// Mitsubishi GX Works2 project: SEMICON_SORTER_ENV   PLC: FX3U/FX3UC

PROGRAM MAIN
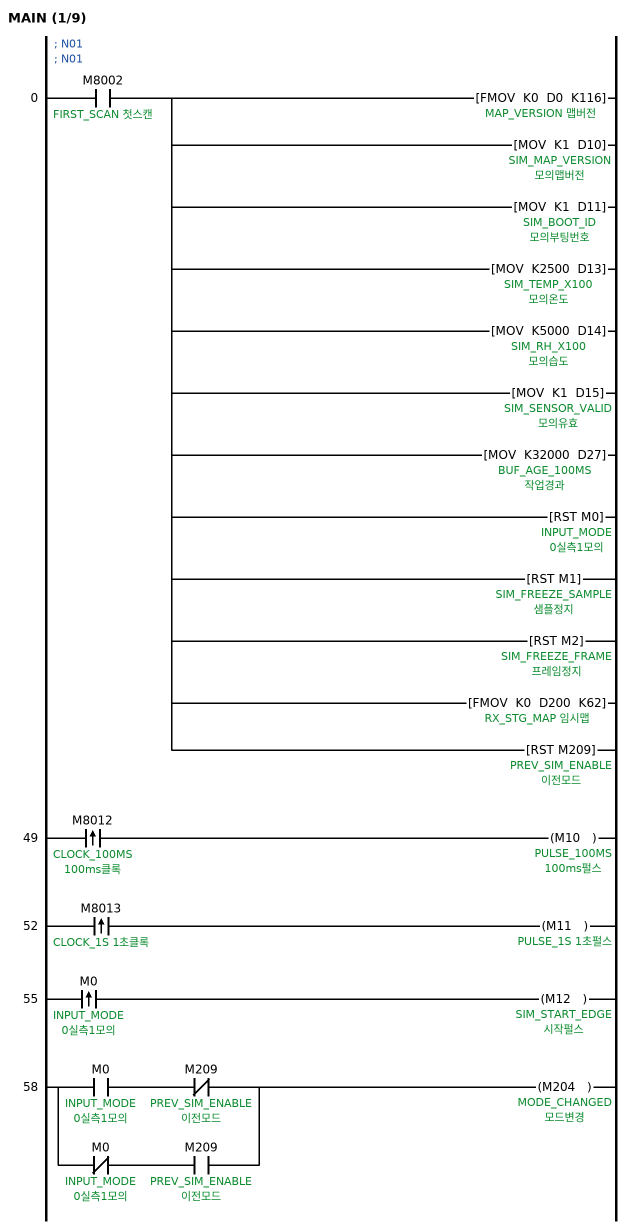
; 
; N01
; N01
0     LD      M8002  ; FIRST_SCAN 첫스캔
      FMOV    K0 D0 K116  ; MAP_VERSION 맵버전
      MOV     K1 D10  ; SIM_MAP_VERSION 모의맵버전
      MOV     K1 D11  ; SIM_BOOT_ID 모의부팅번호
      MOV     K2500 D13  ; SIM_TEMP_X100 모의온도
      MOV     K5000 D14  ; SIM_RH_X100 모의습도
      MOV     K1 D15  ; SIM_SENSOR_VALID 모의유효
      MOV     K32000 D27  ; BUF_AGE_100MS 작업경과
      RST     M0  ; INPUT_MODE 0실측1모의
      RST     M1  ; SIM_FREEZE_SAMPLE 샘플정지
      RST     M2  ; SIM_FREEZE_FRAME 프레임정지
      FMOV    K0 D200 K62  ; RX_STG_MAP 임시맵
      RST     M209  ; PREV_SIM_ENABLE 이전모드
49    LDP     M8012  ; CLOCK_100MS 100ms클록
      OUT     M10  ; PULSE_100MS 100ms펄스
52    LDP     M8013  ; CLOCK_1S 1초클록
      OUT     M11  ; PULSE_1S 1초펄스
55    LDP     M0  ; INPUT_MODE 0실측1모의
      OUT     M12  ; SIM_START_EDGE 시작펄스
58    LD      M0  ; INPUT_MODE 0실측1모의
      ANI     M209  ; PREV_SIM_ENABLE 이전모드
      LDI     M0  ; INPUT_MODE 0실측1모의
      AND     M209  ; PREV_SIM_ENABLE 이전모드
      ORB
      OUT     M204  ; MODE_CHANGED 모드변경
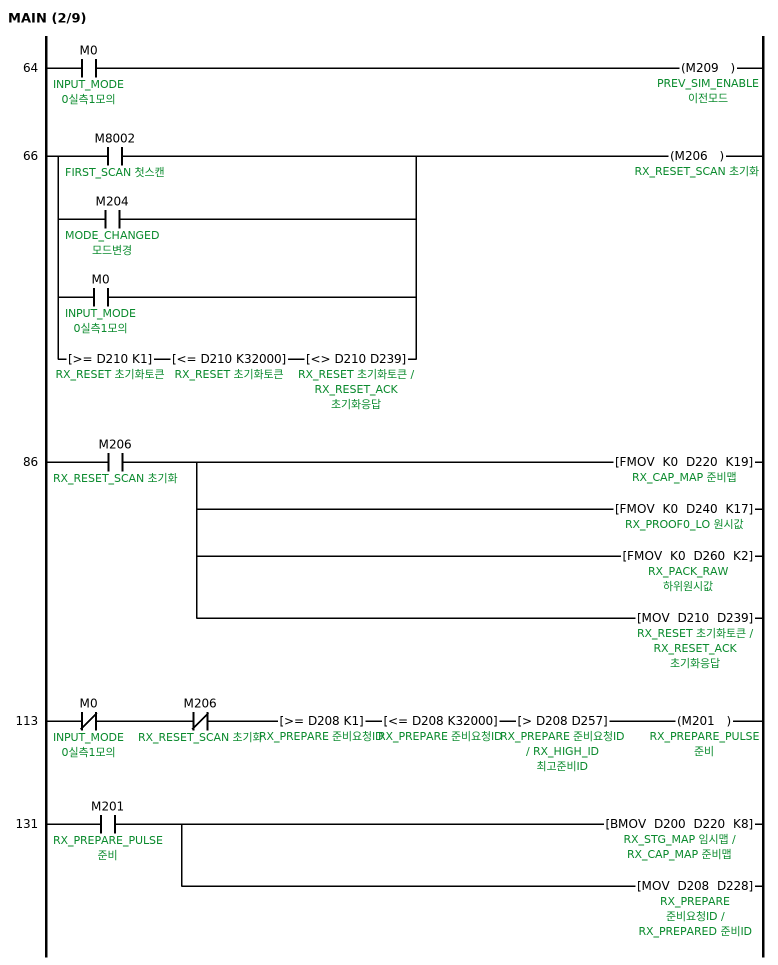
64    LD      M0  ; INPUT_MODE 0실측1모의
      OUT     M209  ; PREV_SIM_ENABLE 이전모드
66    LD      M8002  ; FIRST_SCAN 첫스캔
      OR      M204  ; MODE_CHANGED 모드변경
      OR      M0  ; INPUT_MODE 0실측1모의
      LD>=    D210 K1  ; RX_RESET 초기화토큰
      AND<=   D210 K32000  ; RX_RESET 초기화토큰
      AND<>   D210 D239  ; RX_RESET 초기화토큰 / RX_RESET_ACK 초기화응답
      ORB
      OUT     M206  ; RX_RESET_SCAN 초기화
86    LD      M206  ; RX_RESET_SCAN 초기화
      FMOV    K0 D220 K19  ; RX_CAP_MAP 준비맵
      FMOV    K0 D240 K17  ; RX_PROOF0_LO 원시값
      FMOV    K0 D260 K2  ; RX_PACK_RAW 하위원시값
      MOV     D210 D239
113   LDI     M0  ; INPUT_MODE 0실측1모의
      ANI     M206  ; RX_RESET_SCAN 초기화
      AND>=   D208 K1  ; RX_PREPARE 준비요청ID
      AND<=   D208 K32000  ; RX_PREPARE 준비요청ID
      AND>    D208 D257  ; RX_PREPARE 준비요청ID / RX_HIGH_ID 최고준비ID
      OUT     M201  ; RX_PREPARE_PULSE 준비
131   LD      M201  ; RX_PREPARE_PULSE 준비
      BMOV    D200 D220 K8
      MOV     D208 D228  ; RX_PREPARED 준비ID
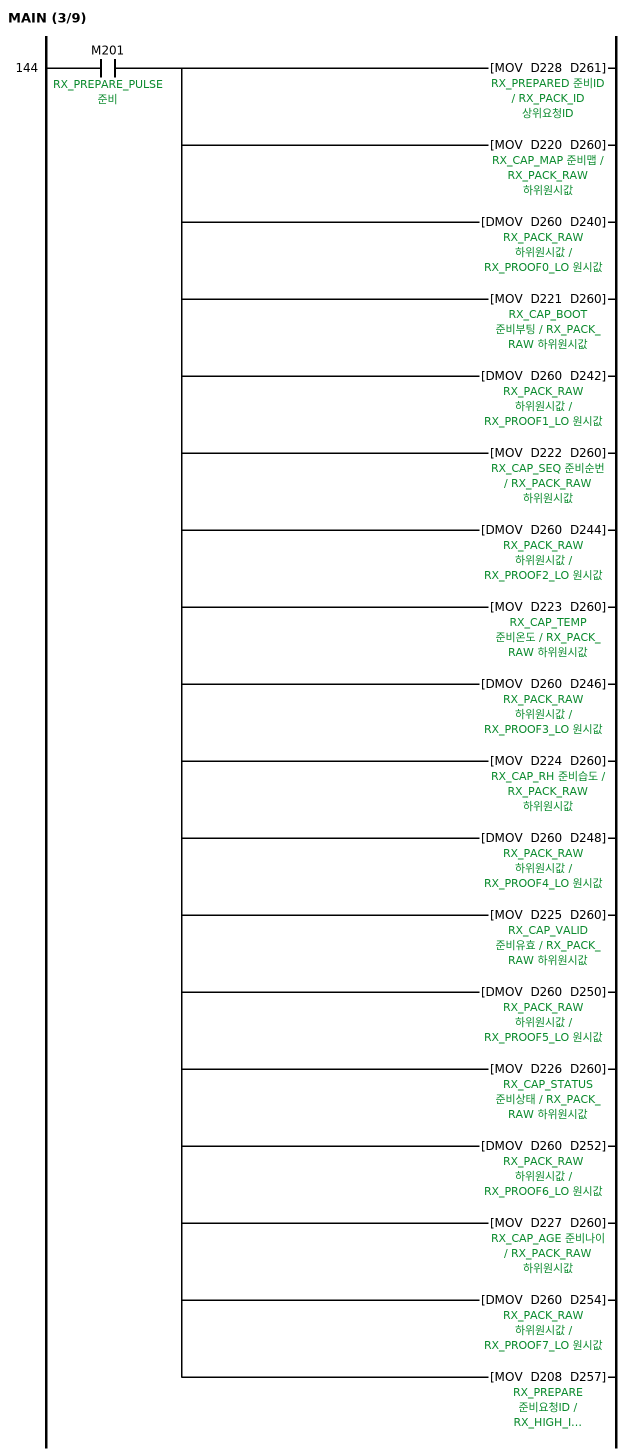
144   LD      M201  ; RX_PREPARE_PULSE 준비
      MOV     D228 D261  ; RX_PACK_ID 상위요청ID
      MOV     D220 D260
      DMOV    D260 D240
      MOV     D221 D260  ; RX_CAP_BOOT 준비부팅
      DMOV    D260 D242  ; RX_PROOF1_LO 원시값
      MOV     D222 D260  ; RX_CAP_SEQ 준비순번
      DMOV    D260 D244  ; RX_PROOF2_LO 원시값
      MOV     D223 D260  ; RX_CAP_TEMP 준비온도
      DMOV    D260 D246  ; RX_PROOF3_LO 원시값
      MOV     D224 D260  ; RX_CAP_RH 준비습도
      DMOV    D260 D248  ; RX_PROOF4_LO 원시값
      MOV     D225 D260  ; RX_CAP_VALID 준비유효
      DMOV    D260 D250  ; RX_PROOF5_LO 원시값
      MOV     D226 D260  ; RX_CAP_STATUS 준비상태
      DMOV    D260 D252  ; RX_PROOF6_LO 원시값
      MOV     D227 D260  ; RX_CAP_AGE 준비나이
      DMOV    D260 D254  ; RX_PROOF7_LO 원시값
      MOV     D208 D257
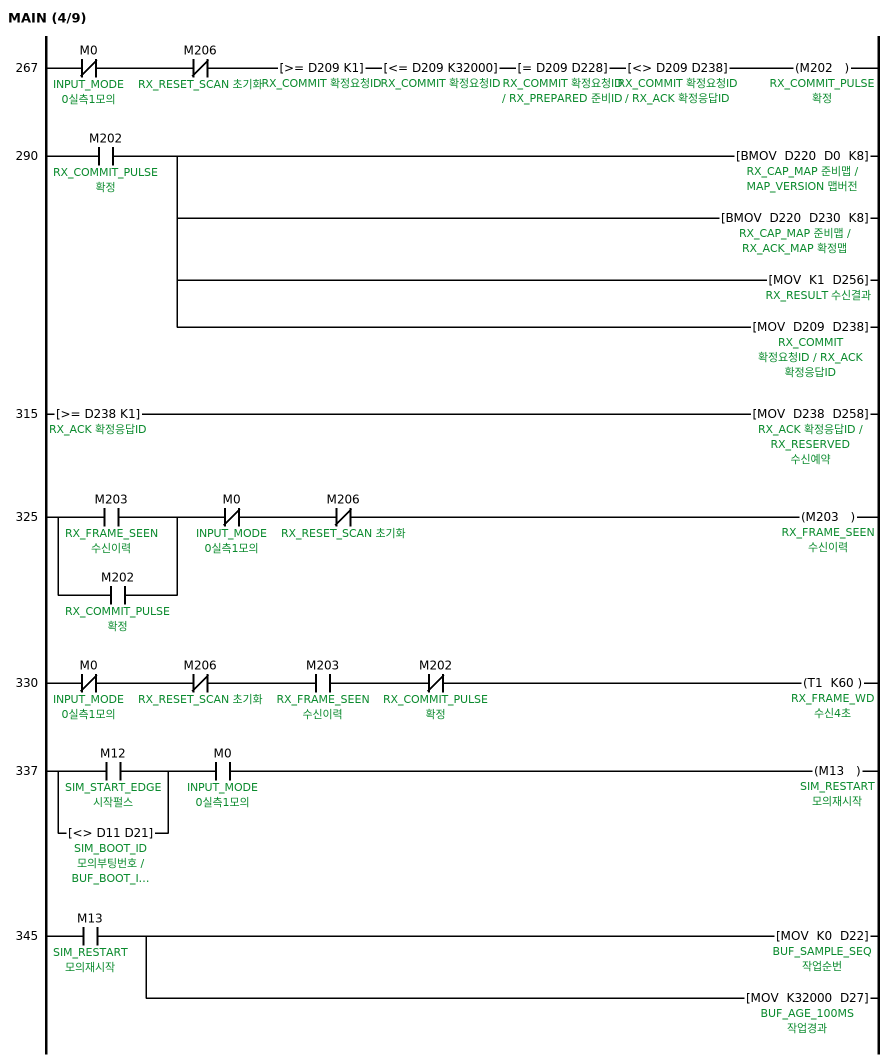
267   LDI     M0  ; INPUT_MODE 0실측1모의
      ANI     M206  ; RX_RESET_SCAN 초기화
      AND>=   D209 K1  ; RX_COMMIT 확정요청ID
      AND<=   D209 K32000  ; RX_COMMIT 확정요청ID
      AND=    D209 D228  ; RX_COMMIT 확정요청ID / RX_PREPARED 준비ID
      AND<>   D209 D238  ; RX_COMMIT 확정요청ID / RX_ACK 확정응답ID
      OUT     M202  ; RX_COMMIT_PULSE 확정
290   LD      M202  ; RX_COMMIT_PULSE 확정
      BMOV    D220 D0 K8
      BMOV    D220 D230 K8  ; RX_ACK_MAP 확정맵
      MOV     K1 D256  ; RX_RESULT 수신결과
      MOV     D209 D238
315   LD>=    D238 K1  ; RX_ACK 확정응답ID
      MOV     D238 D258  ; RX_RESERVED 수신예약
325   LD      M203  ; RX_FRAME_SEEN 수신이력
      OR      M202  ; RX_COMMIT_PULSE 확정
      ANI     M0  ; INPUT_MODE 0실측1모의
      ANI     M206  ; RX_RESET_SCAN 초기화
      OUT     M203  ; RX_FRAME_SEEN 수신이력
330   LDI     M0  ; INPUT_MODE 0실측1모의
      ANI     M206  ; RX_RESET_SCAN 초기화
      AND     M203  ; RX_FRAME_SEEN 수신이력
      ANI     M202  ; RX_COMMIT_PULSE 확정
      OUT     T1 K60  ; RX_FRAME_WD 수신4초
337   LD      M12  ; SIM_START_EDGE 시작펄스
      OR<>    D11 D21  ; SIM_BOOT_ID 모의부팅번호 / BUF_BOOT_ID 작업부팅번호
      AND     M0  ; INPUT_MODE 0실측1모의
      OUT     M13  ; SIM_RESTART 모의재시작
345   LD      M13  ; SIM_RESTART 모의재시작
      MOV     K0 D22  ; BUF_SAMPLE_SEQ 작업순번
      MOV     K32000 D27
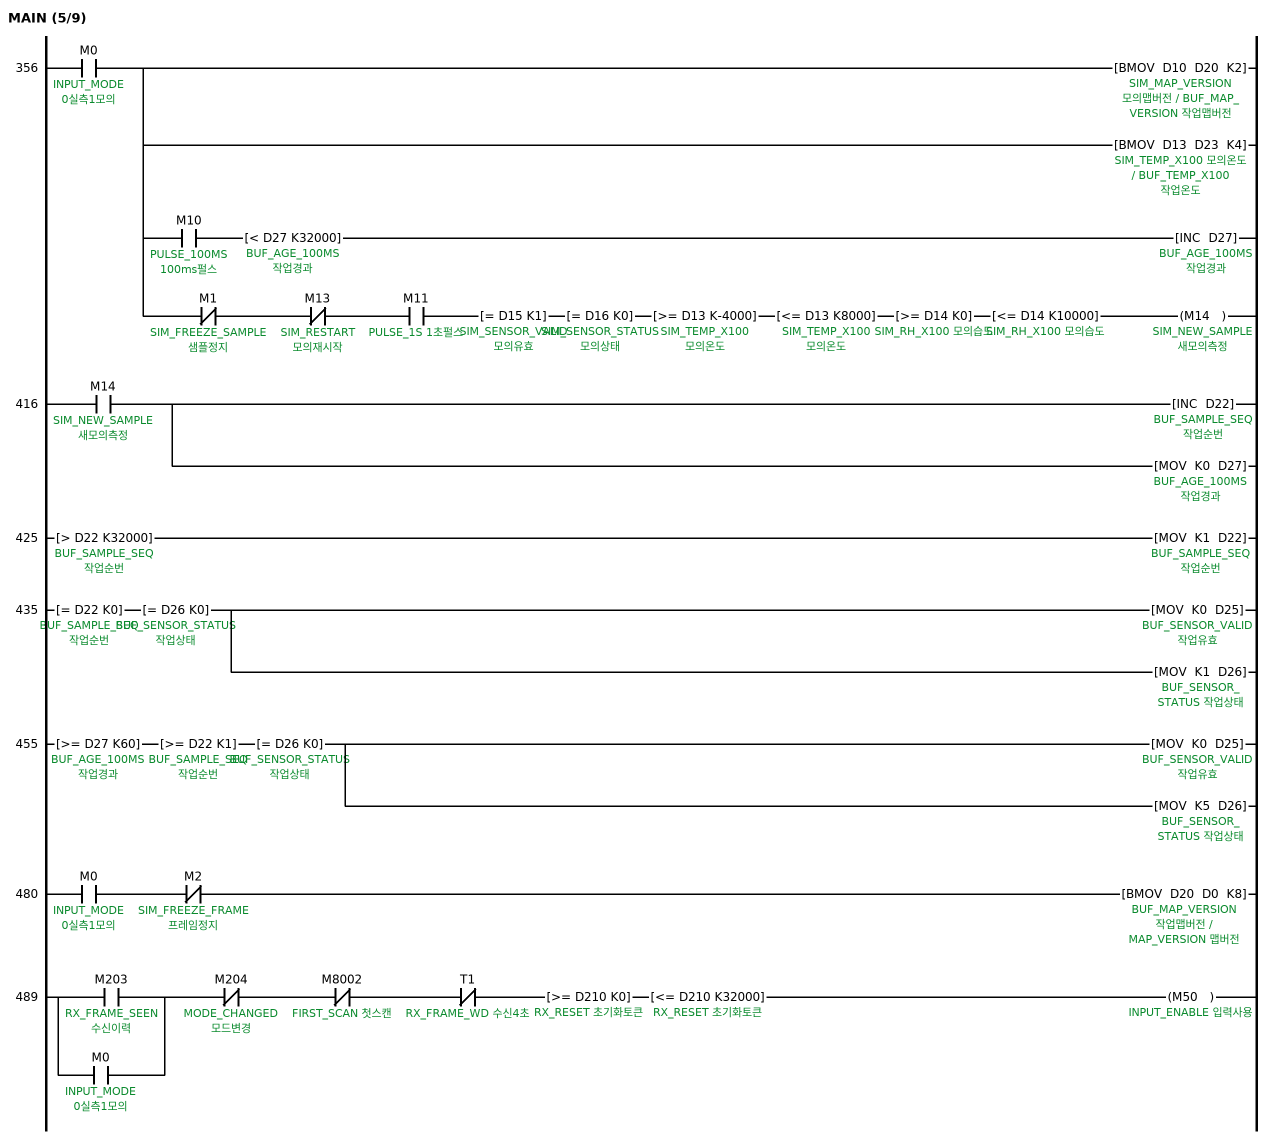
356   LD      M0  ; INPUT_MODE 0실측1모의
      BMOV    D10 D20 K2  ; BUF_MAP_VERSION 작업맵버전
      BMOV    D13 D23 K4  ; BUF_TEMP_X100 작업온도
      MPS
      AND     M10  ; PULSE_100MS 100ms펄스
      AND<    D27 K32000  ; BUF_AGE_100MS 작업경과
      INC     D27
      MPP
      ANI     M1  ; SIM_FREEZE_SAMPLE 샘플정지
      ANI     M13  ; SIM_RESTART 모의재시작
      AND     M11  ; PULSE_1S 1초펄스
      AND=    D15 K1  ; SIM_SENSOR_VALID 모의유효
      AND=    D16 K0  ; SIM_SENSOR_STATUS 모의상태
      AND>=   D13 K-4000  ; SIM_TEMP_X100 모의온도
      AND<=   D13 K8000  ; SIM_TEMP_X100 모의온도
      AND>=   D14 K0  ; SIM_RH_X100 모의습도
      AND<=   D14 K10000  ; SIM_RH_X100 모의습도
      OUT     M14  ; SIM_NEW_SAMPLE 새모의측정
416   LD      M14  ; SIM_NEW_SAMPLE 새모의측정
      INC     D22
      MOV     K0 D27
425   LD>     D22 K32000  ; BUF_SAMPLE_SEQ 작업순번
      MOV     K1 D22
435   LD=     D22 K0  ; BUF_SAMPLE_SEQ 작업순번
      AND=    D26 K0  ; BUF_SENSOR_STATUS 작업상태
      MOV     K0 D25  ; BUF_SENSOR_VALID 작업유효
      MOV     K1 D26
455   LD>=    D27 K60  ; BUF_AGE_100MS 작업경과
      AND>=   D22 K1  ; BUF_SAMPLE_SEQ 작업순번
      AND=    D26 K0  ; BUF_SENSOR_STATUS 작업상태
      MOV     K0 D25
      MOV     K5 D26
480   LD      M0  ; INPUT_MODE 0실측1모의
      ANI     M2  ; SIM_FREEZE_FRAME 프레임정지
      BMOV    D20 D0 K8
489   LD      M203  ; RX_FRAME_SEEN 수신이력
      OR      M0  ; INPUT_MODE 0실측1모의
      ANI     M204  ; MODE_CHANGED 모드변경
      ANI     M8002  ; FIRST_SCAN 첫스캔
      ANI     T1  ; RX_FRAME_WD 수신4초
      AND>=   D210 K0  ; RX_RESET 초기화토큰
      AND<=   D210 K32000  ; RX_RESET 초기화토큰
      OUT     M50  ; INPUT_ENABLE 입력사용
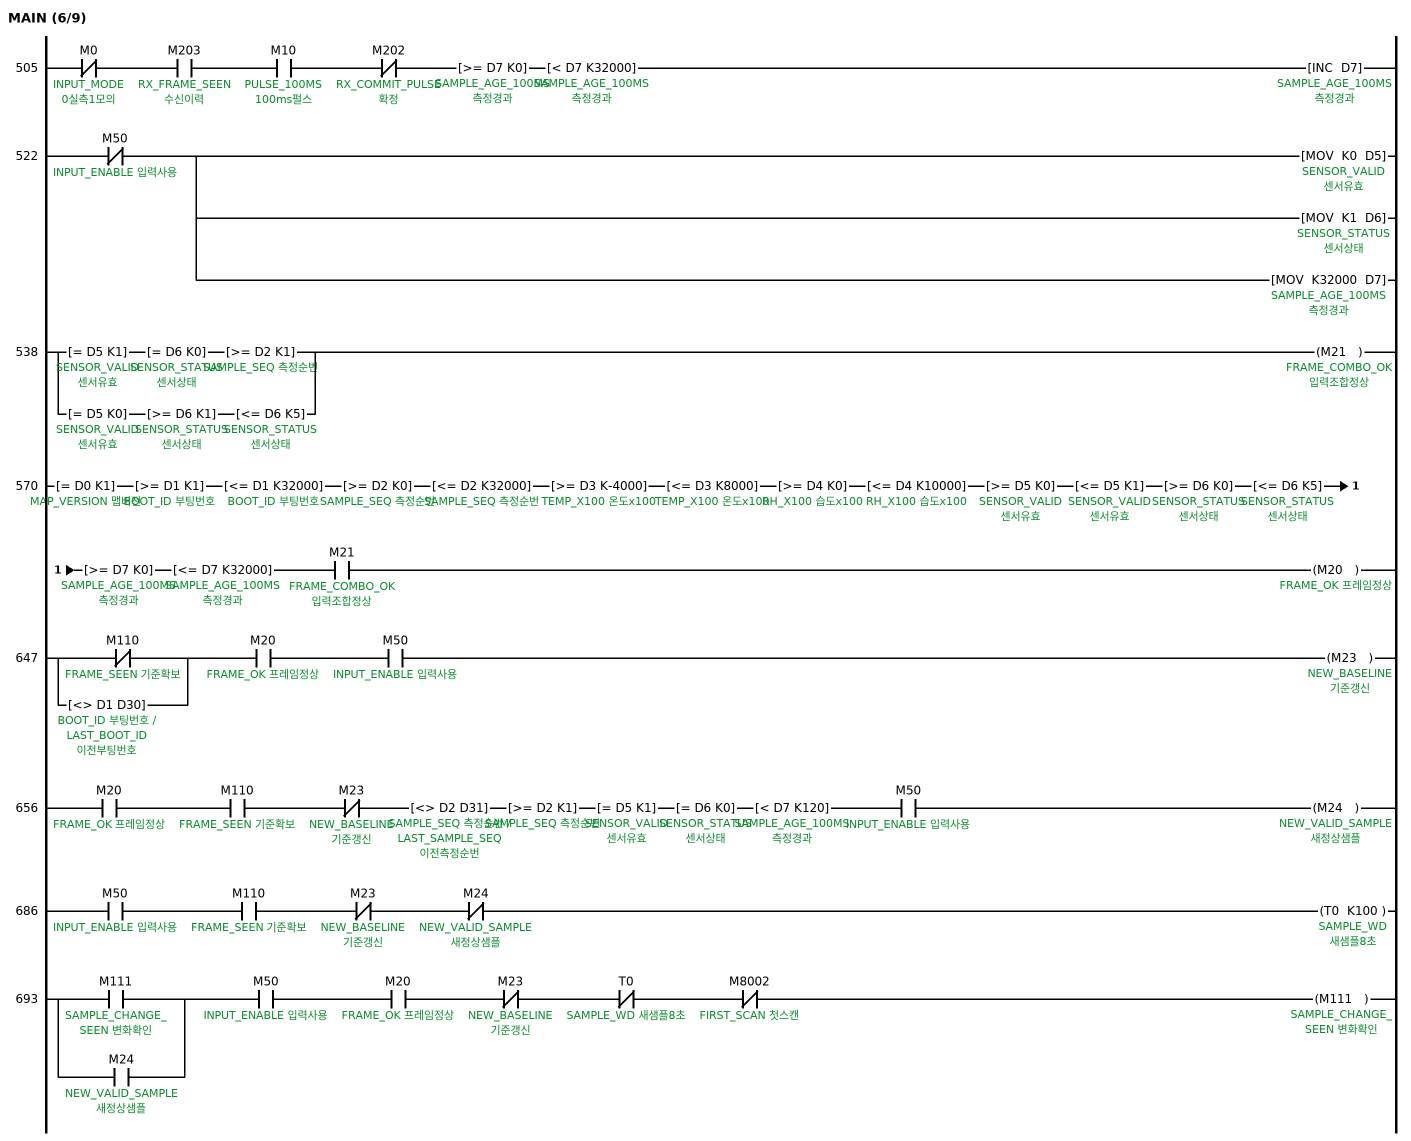
505   LDI     M0  ; INPUT_MODE 0실측1모의
      AND     M203  ; RX_FRAME_SEEN 수신이력
      AND     M10  ; PULSE_100MS 100ms펄스
      ANI     M202  ; RX_COMMIT_PULSE 확정
      AND>=   D7 K0  ; SAMPLE_AGE_100MS 측정경과
      AND<    D7 K32000  ; SAMPLE_AGE_100MS 측정경과
      INC     D7
522   LDI     M50  ; INPUT_ENABLE 입력사용
      MOV     K0 D5  ; SENSOR_VALID 센서유효
      MOV     K1 D6  ; SENSOR_STATUS 센서상태
      MOV     K32000 D7
538   LD=     D5 K1  ; SENSOR_VALID 센서유효
      AND=    D6 K0  ; SENSOR_STATUS 센서상태
      AND>=   D2 K1  ; SAMPLE_SEQ 측정순번
      LD=     D5 K0  ; SENSOR_VALID 센서유효
      AND>=   D6 K1  ; SENSOR_STATUS 센서상태
      AND<=   D6 K5  ; SENSOR_STATUS 센서상태
      ORB
      OUT     M21  ; FRAME_COMBO_OK 입력조합정상
570   LD=     D0 K1  ; MAP_VERSION 맵버전
      AND>=   D1 K1  ; BOOT_ID 부팅번호
      AND<=   D1 K32000  ; BOOT_ID 부팅번호
      AND>=   D2 K0  ; SAMPLE_SEQ 측정순번
      AND<=   D2 K32000  ; SAMPLE_SEQ 측정순번
      AND>=   D3 K-4000  ; TEMP_X100 온도x100
      AND<=   D3 K8000  ; TEMP_X100 온도x100
      AND>=   D4 K0  ; RH_X100 습도x100
      AND<=   D4 K10000  ; RH_X100 습도x100
      AND>=   D5 K0  ; SENSOR_VALID 센서유효
      AND<=   D5 K1  ; SENSOR_VALID 센서유효
      AND>=   D6 K0  ; SENSOR_STATUS 센서상태
      AND<=   D6 K5  ; SENSOR_STATUS 센서상태
      AND>=   D7 K0  ; SAMPLE_AGE_100MS 측정경과
      AND<=   D7 K32000  ; SAMPLE_AGE_100MS 측정경과
      AND     M21  ; FRAME_COMBO_OK 입력조합정상
      OUT     M20  ; FRAME_OK 프레임정상
647   LDI     M110  ; FRAME_SEEN 기준확보
      OR<>    D1 D30  ; BOOT_ID 부팅번호 / LAST_BOOT_ID 이전부팅번호
      AND     M20  ; FRAME_OK 프레임정상
      AND     M50  ; INPUT_ENABLE 입력사용
      OUT     M23  ; NEW_BASELINE 기준갱신
656   LD      M20  ; FRAME_OK 프레임정상
      AND     M110  ; FRAME_SEEN 기준확보
      ANI     M23  ; NEW_BASELINE 기준갱신
      AND<>   D2 D31  ; SAMPLE_SEQ 측정순번 / LAST_SAMPLE_SEQ 이전측정순번
      AND>=   D2 K1  ; SAMPLE_SEQ 측정순번
      AND=    D5 K1  ; SENSOR_VALID 센서유효
      AND=    D6 K0  ; SENSOR_STATUS 센서상태
      AND<    D7 K120  ; SAMPLE_AGE_100MS 측정경과
      AND     M50  ; INPUT_ENABLE 입력사용
      OUT     M24  ; NEW_VALID_SAMPLE 새정상샘플
686   LD      M50  ; INPUT_ENABLE 입력사용
      AND     M110  ; FRAME_SEEN 기준확보
      ANI     M23  ; NEW_BASELINE 기준갱신
      ANI     M24  ; NEW_VALID_SAMPLE 새정상샘플
      OUT     T0 K100  ; SAMPLE_WD 새샘플8초
693   LD      M111  ; SAMPLE_CHANGE_SEEN 변화확인
      OR      M24  ; NEW_VALID_SAMPLE 새정상샘플
      AND     M50  ; INPUT_ENABLE 입력사용
      AND     M20  ; FRAME_OK 프레임정상
      ANI     M23  ; NEW_BASELINE 기준갱신
      ANI     T0  ; SAMPLE_WD 새샘플8초
      ANI     M8002  ; FIRST_SCAN 첫스캔
      OUT     M111  ; SAMPLE_CHANGE_SEEN 변화확인
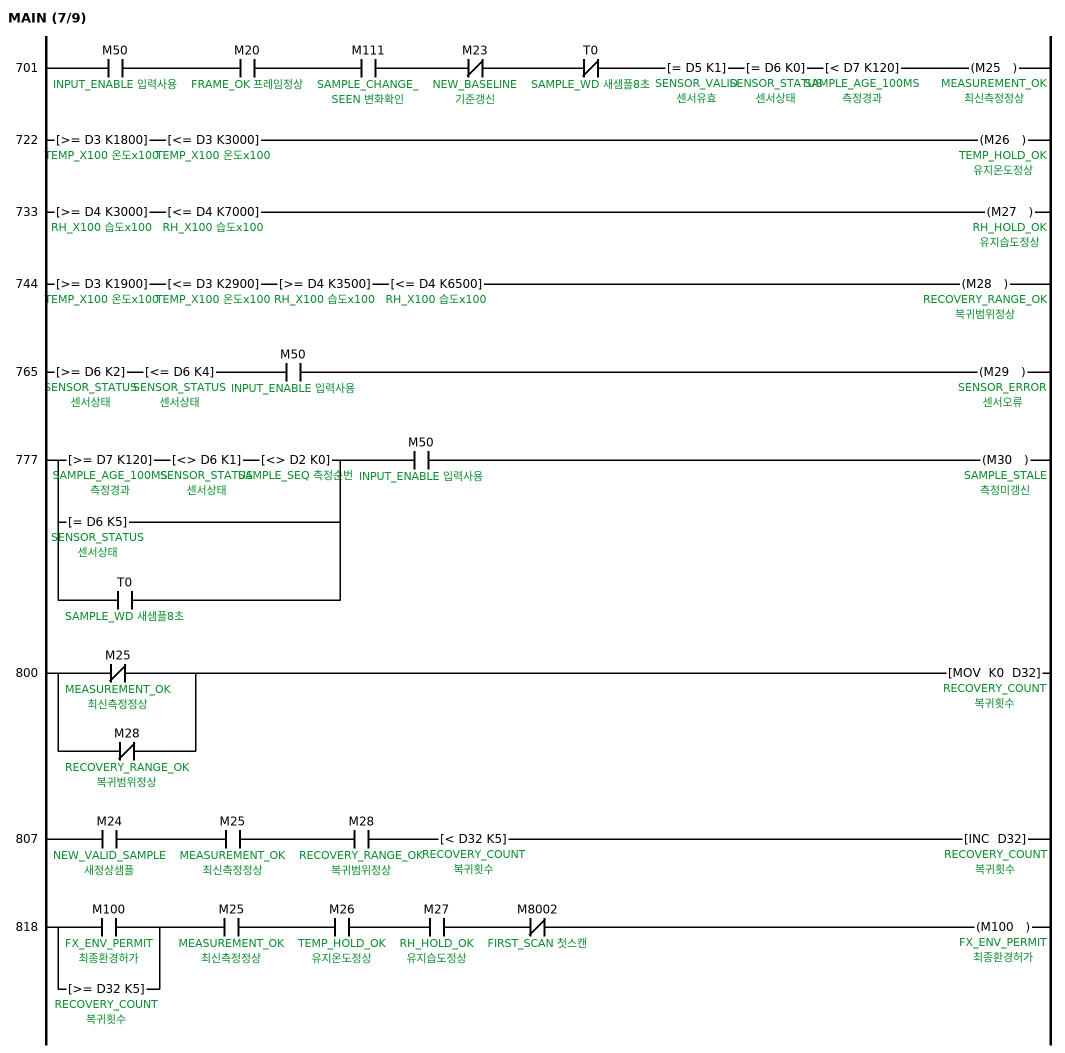
701   LD      M50  ; INPUT_ENABLE 입력사용
      AND     M20  ; FRAME_OK 프레임정상
      AND     M111  ; SAMPLE_CHANGE_SEEN 변화확인
      ANI     M23  ; NEW_BASELINE 기준갱신
      ANI     T0  ; SAMPLE_WD 새샘플8초
      AND=    D5 K1  ; SENSOR_VALID 센서유효
      AND=    D6 K0  ; SENSOR_STATUS 센서상태
      AND<    D7 K120  ; SAMPLE_AGE_100MS 측정경과
      OUT     M25  ; MEASUREMENT_OK 최신측정정상
722   LD>=    D3 K1800  ; TEMP_X100 온도x100
      AND<=   D3 K3000  ; TEMP_X100 온도x100
      OUT     M26  ; TEMP_HOLD_OK 유지온도정상
733   LD>=    D4 K3000  ; RH_X100 습도x100
      AND<=   D4 K7000  ; RH_X100 습도x100
      OUT     M27  ; RH_HOLD_OK 유지습도정상
744   LD>=    D3 K1900  ; TEMP_X100 온도x100
      AND<=   D3 K2900  ; TEMP_X100 온도x100
      AND>=   D4 K3500  ; RH_X100 습도x100
      AND<=   D4 K6500  ; RH_X100 습도x100
      OUT     M28  ; RECOVERY_RANGE_OK 복귀범위정상
765   LD>=    D6 K2  ; SENSOR_STATUS 센서상태
      AND<=   D6 K4  ; SENSOR_STATUS 센서상태
      AND     M50  ; INPUT_ENABLE 입력사용
      OUT     M29  ; SENSOR_ERROR 센서오류
777   LD>=    D7 K120  ; SAMPLE_AGE_100MS 측정경과
      AND<>   D6 K1  ; SENSOR_STATUS 센서상태
      AND<>   D2 K0  ; SAMPLE_SEQ 측정순번
      OR=     D6 K5  ; SENSOR_STATUS 센서상태
      OR      T0  ; SAMPLE_WD 새샘플8초
      AND     M50  ; INPUT_ENABLE 입력사용
      OUT     M30  ; SAMPLE_STALE 측정미갱신
800   LDI     M25  ; MEASUREMENT_OK 최신측정정상
      ORI     M28  ; RECOVERY_RANGE_OK 복귀범위정상
      MOV     K0 D32  ; RECOVERY_COUNT 복귀횟수
807   LD      M24  ; NEW_VALID_SAMPLE 새정상샘플
      AND     M25  ; MEASUREMENT_OK 최신측정정상
      AND     M28  ; RECOVERY_RANGE_OK 복귀범위정상
      AND<    D32 K5  ; RECOVERY_COUNT 복귀횟수
      INC     D32
818   LD      M100  ; FX_ENV_PERMIT 최종환경허가
      OR>=    D32 K5  ; RECOVERY_COUNT 복귀횟수
      AND     M25  ; MEASUREMENT_OK 최신측정정상
      AND     M26  ; TEMP_HOLD_OK 유지온도정상
      AND     M27  ; RH_HOLD_OK 유지습도정상
      ANI     M8002  ; FIRST_SCAN 첫스캔
      OUT     M100  ; FX_ENV_PERMIT 최종환경허가
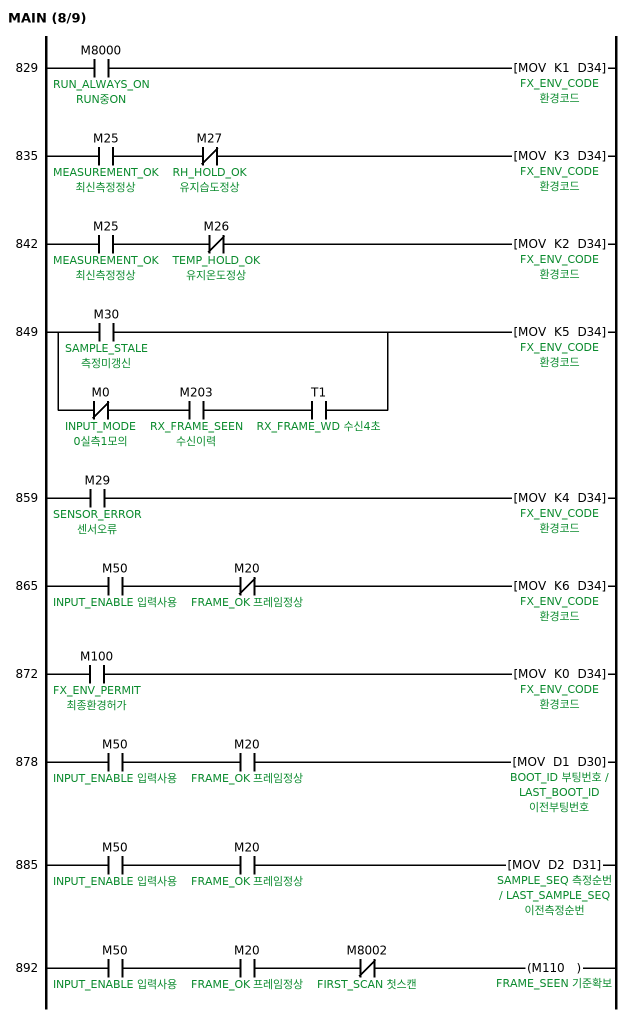
829   LD      M8000  ; RUN_ALWAYS_ON RUN중ON
      MOV     K1 D34  ; FX_ENV_CODE 환경코드
835   LD      M25  ; MEASUREMENT_OK 최신측정정상
      ANI     M27  ; RH_HOLD_OK 유지습도정상
      MOV     K3 D34
842   LD      M25  ; MEASUREMENT_OK 최신측정정상
      ANI     M26  ; TEMP_HOLD_OK 유지온도정상
      MOV     K2 D34
849   LD      M30  ; SAMPLE_STALE 측정미갱신
      LDI     M0  ; INPUT_MODE 0실측1모의
      AND     M203  ; RX_FRAME_SEEN 수신이력
      AND     T1  ; RX_FRAME_WD 수신4초
      ORB
      MOV     K5 D34
859   LD      M29  ; SENSOR_ERROR 센서오류
      MOV     K4 D34
865   LD      M50  ; INPUT_ENABLE 입력사용
      ANI     M20  ; FRAME_OK 프레임정상
      MOV     K6 D34
872   LD      M100  ; FX_ENV_PERMIT 최종환경허가
      MOV     K0 D34
878   LD      M50  ; INPUT_ENABLE 입력사용
      AND     M20  ; FRAME_OK 프레임정상
      MOV     D1 D30
885   LD      M50  ; INPUT_ENABLE 입력사용
      AND     M20  ; FRAME_OK 프레임정상
      MOV     D2 D31
892   LD      M50  ; INPUT_ENABLE 입력사용
      AND     M20  ; FRAME_OK 프레임정상
      ANI     M8002  ; FIRST_SCAN 첫스캔
      OUT     M110  ; FRAME_SEEN 기준확보
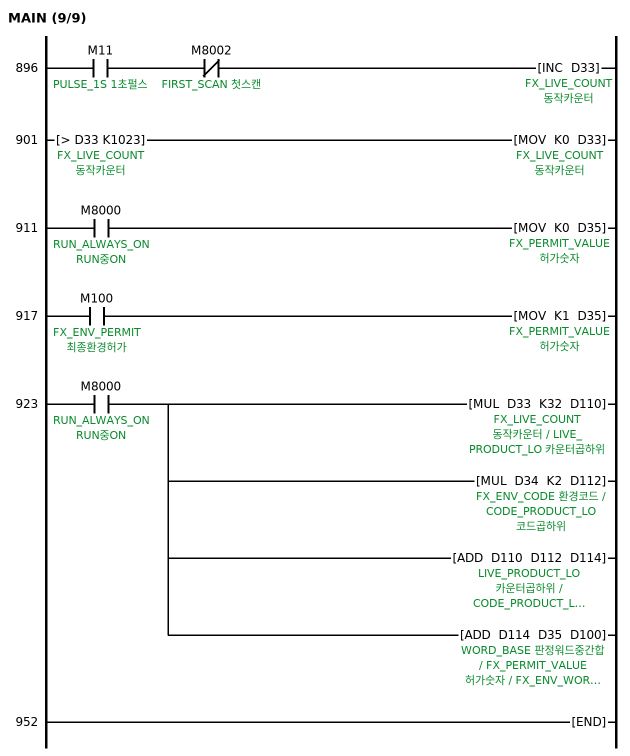
896   LD      M11  ; PULSE_1S 1초펄스
      ANI     M8002  ; FIRST_SCAN 첫스캔
      INC     D33  ; FX_LIVE_COUNT 동작카운터
901   LD>     D33 K1023  ; FX_LIVE_COUNT 동작카운터
      MOV     K0 D33
911   LD      M8000  ; RUN_ALWAYS_ON RUN중ON
      MOV     K0 D35  ; FX_PERMIT_VALUE 허가숫자
917   LD      M100  ; FX_ENV_PERMIT 최종환경허가
      MOV     K1 D35
923   LD      M8000  ; RUN_ALWAYS_ON RUN중ON
      MUL     D33 K32 D110  ; LIVE_PRODUCT_LO 카운터곱하위
      MUL     D34 K2 D112  ; CODE_PRODUCT_LO 코드곱하위
      ADD     D110 D112 D114  ; WORD_BASE 판정워드중간합
      ADD     D114 D35 D100  ; FX_ENV_WORD 최종판정워드
952   END
END_PROGRAM

// device comments not shown above
D24  ; BUF_RH_X100 작업습도
D111  ; LIVE_PRODUCT_HI 카운터곱상위
D113  ; CODE_PRODUCT_HI 코드곱상위
D115  ; RESERVED 예약미사용
D201  ; RX_STG_BOOT 임시부팅
D202  ; RX_STG_SEQ 임시순번
D203  ; RX_STG_TEMP 임시온도
D204  ; RX_STG_RH 임시습도
D205  ; RX_STG_VALID 임시유효
D206  ; RX_STG_STATUS 임시상태
D207  ; RX_STG_AGE 임시나이
D231  ; RX_ACK_BOOT 확정부팅
D232  ; RX_ACK_SEQ 확정순번
D233  ; RX_ACK_TEMP 확정온도
D234  ; RX_ACK_RH 확정습도
D235  ; RX_ACK_VALID 확정유효
D236  ; RX_ACK_STATUS 확정상태
D237  ; RX_ACK_AGE 확정나이
D241  ; RX_PROOF0_HI 준비ID
D243  ; RX_PROOF1_HI 준비ID
D245  ; RX_PROOF2_HI 준비ID
D247  ; RX_PROOF3_HI 준비ID
D249  ; RX_PROOF4_HI 준비ID
D251  ; RX_PROOF5_HI 준비ID
D253  ; RX_PROOF6_HI 준비ID
D255  ; RX_PROOF7_HI 준비ID
